ABB RAPID module: CalibData.mod

MODULE CalibData
    PERS tooldata punta:=[TRUE,[[24,0,172],[0.945519,0,0.325568,0]],[0.1,[0,0,1],[1,0,0,0],0,0,0]];
    TASK PERS wobjdata WOCaja:=[FALSE,TRUE,"",[[253.5,-72.5,200],[0,0.707107,0.707107,0]],[[0,0,0],[1,0,0,0]]];
ENDMODULE
